FUNCTION_BLOCK F (* Negative C4: the same dispatch written as separate IFs in a shared algorithm *)
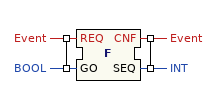
  EVENT_INPUT
    REQ WITH GO;
  END_EVENT
  EVENT_OUTPUT
    CNF WITH SEQ;
  END_EVENT
  VAR_INPUT
    GO : BOOL;
  END_VAR
  VAR_OUTPUT
    SEQ : INT;
  END_VAR
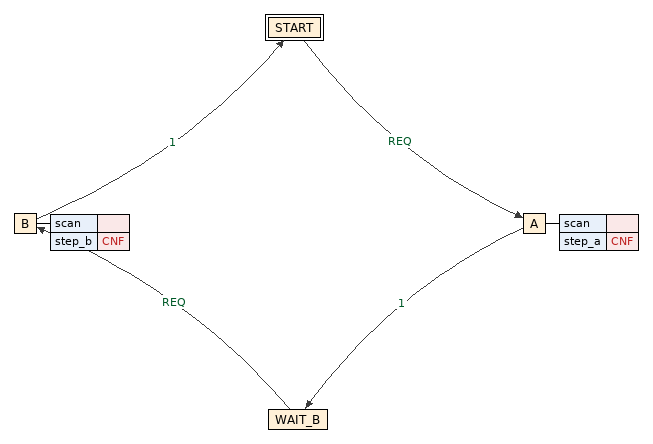
  EC_STATES
    START;
    A : scan, step_a -> CNF;
    WAIT_B;
    B : scan, step_b -> CNF;
  END_STATES
  EC_TRANSITIONS
    START TO A := REQ;
    A TO WAIT_B := 1;
    WAIT_B TO B := REQ;
    B TO START := 1;
  END_TRANSITIONS
  ALGORITHM scan IN ST:
IF SEQ = 0 THEN
  SEQ := 1;
END_IF;
IF SEQ = 1 THEN
  SEQ := 0;
END_IF;
  END_ALGORITHM
  ALGORITHM step_a IN ST:
SEQ := 0;
IF GO THEN
  SEQ := 1;
END_IF;
  END_ALGORITHM
  ALGORITHM step_b IN ST:
IF NOT GO THEN
  SEQ := 0;
END_IF;
  END_ALGORITHM
END_FUNCTION_BLOCK
